TYPE ST_Nidec :
STRUCT
	StatusWord     AT %I* : WORD;     // Input from Receive PDO Mapping 6
	ControlWord     AT %Q* : WORD;      // Output to Transmit PDO Mapping 6
	
	actVelocity AT %I*: INT;
	targetVelocity AT %Q*: INT;
END_STRUCT
END_TYPE

(* stored: Version 1.1.0.1, ProductVersion 3.1.4024.12
   DUT ST_Nidec: Id {4a038cd4-9b62-4041-9ddf-9d5b9b94b29b} *)
